KUKA KRL program: Section1.src

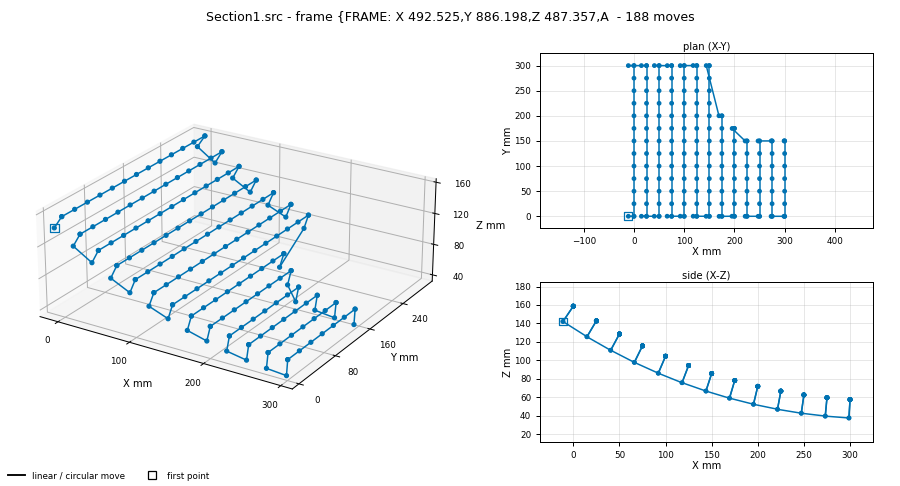
[picture p0: tool path of Section1.src in frame {FRAME: X 492.525,Y 886.198,Z 487.357,A , 188 of 189 moves have a stored position in this frame; points joined in program order, loops and branches not executed]
&ACCESS RVP
&REL 1
&PARAM TEMPLATE = C:\KRC\Roboter\Template\vorgabe
&PARAM EDITMASK = *
DEF Section1 ( )
EXT BAS (BAS_COMMAND :IN,REAL :IN )


; GLOBAL INTERRUPT DECL 3 WHEN $STOPMESS==TRUE DO IR_STOPM ( )
; INTERRUPT ON 3

;FOLD Initialise and set default speed
BAS (#INITMOV,0)
BAS (#VEL_PTP,100)
BAS (#ACC_PTP,20)
$VEL.CP=0.2
BAS (#TOOL,0)
BAS (#BASE,0)
;ENDFOLD

;;FOLD STARTPOS
;$BWDSTART = FALSE
;PDAT_ACT = PDEFAULT
;BAS(#PTP_DAT)
;FDAT_ACT = {TOOL_NO 0,BASE_NO 0,IPO_FRAME #BASE}
;BAS(#FRAMES)
;;ENDFOLD

$ADVANCE = 5

;FOLD ---- Quickly skip BCO ----
; PTP $AXIS_ACT
;ENDFOLD

;FOLD ---- GO HOME ----
; PTP {A1 0.000, A2 -90.000, A3 90.000, A4 0.000, A5 0.000, A6 0.000, E1 0, E2 0, E3 0, E4 0, E5 0, E6 0}
;ENDFOLD


; Program generated by VerticalBot Studio for KUKA KR 5 arc on 25/10/2026 12:00:00
; Using nominal kinematics.
; ---- Setting reference (Base) ----
; BASE_DATA[1] = {FRAME: X 492.525,Y 886.198,Z 487.357,A 87.824,B 90.000,C 0.000}
$BASE = {FRAME: X 492.525,Y 886.198,Z 487.357,A 87.824,B 90.000,C 0.000}
; $BASE = BASE_DATA[1]
; --------------------------
; ---- Setting tool (TCP) ----
$TOOL = {FRAME: X 25.000,Y 0.000,Z 225.000,A 0.000,B 30.000,C 0.000}
; --------------------------
; show Paint gun
$VEL.CP = 1.00000
PTP {A1 -66.38630,A2 -78.06180,A3 119.38400,A4 136.02800,A5 16.79140,A6 145.96200}
LIN {X -11.194,Y -0.005,Z 142.140,A 88.999,B 0.694,C 34.030}
LIN {X 0.000,Y 0.000,Z 158.714,A 88.999,B 0.694,C 34.030}
LIN {X 0.000,Y 0.000,Z 158.714,A 88.999,B 0.694,C 34.030}
$VEL.CP = 0.02000
LIN {X 0.000,Y 25.000,Z 158.706,A 88.999,B 0.694,C 34.030}
LIN {X 0.000,Y 50.000,Z 158.698,A 88.999,B 0.694,C 34.030}
LIN {X 0.000,Y 75.000,Z 158.689,A 88.999,B 0.695,C 34.022}
LIN {X 0.000,Y 100.000,Z 158.681,A 88.999,B 0.695,C 34.022}
LIN {X 0.000,Y 125.000,Z 158.672,A 88.999,B 0.695,C 34.022}
LIN {X 0.000,Y 150.000,Z 158.664,A 88.999,B 0.695,C 34.022}
LIN {X 0.000,Y 175.000,Z 158.655,A 88.999,B 0.695,C 34.022}
LIN {X 0.000,Y 200.000,Z 158.647,A 88.999,B 0.695,C 34.022}
LIN {X 0.000,Y 225.000,Z 158.638,A 88.999,B 0.695,C 34.022}
LIN {X 0.000,Y 250.000,Z 158.630,A 88.999,B 0.695,C 34.022}
LIN {X 0.000,Y 275.000,Z 158.628,A 88.985,B 0.696,C 34.438}
LIN {X 0.000,Y 300.000,Z 158.634,A 88.981,B 0.668,C 34.022}
$VEL.CP = 1.00000
LIN {X 0.000,Y 300.000,Z 158.634,A 88.981,B 0.668,C 34.022}
LIN {X -11.192,Y 300.006,Z 142.059,A 88.981,B 0.668,C 34.022}
$VEL.CP = 1.00000
LIN {X 14.800,Y 300.034,Z 125.622,A 88.995,B 0.482,C 30.661}
LIN {X 25.000,Y 300.000,Z 142.825,A 88.995,B 0.482,C 30.661}
LIN {X 25.000,Y 300.000,Z 142.825,A 88.995,B 0.482,C 30.661}
$VEL.CP = 0.02000
LIN {X 25.000,Y 275.000,Z 142.758,A 89.004,B 0.509,C 30.830}
LIN {X 25.000,Y 250.000,Z 142.800,A 89.264,B 0.921,C 30.374}
LIN {X 25.000,Y 225.000,Z 142.817,A 88.955,B 0.414,C 30.654}
LIN {X 25.000,Y 200.000,Z 142.818,A 89.100,B 0.691,C 31.206}
LIN {X 25.000,Y 175.000,Z 142.825,A 88.923,B 0.380,C 30.934}
LIN {X 25.000,Y 150.000,Z 142.711,A 88.930,B 0.392,C 30.935}
LIN {X 25.000,Y 125.000,Z 142.731,A 89.108,B 0.682,C 30.827}
LIN {X 25.000,Y 100.000,Z 142.834,A 88.962,B 0.476,C 31.406}
LIN {X 25.000,Y 75.000,Z 142.753,A 88.812,B 0.195,C 30.940}
LIN {X 25.000,Y 50.000,Z 142.717,A 89.127,B 0.702,C 30.616}
LIN {X 25.000,Y 25.000,Z 142.723,A 89.019,B 0.516,C 30.561}
LIN {X 25.000,Y 0.000,Z 142.733,A 88.984,B 0.455,C 30.523}
$VEL.CP = 1.00000
LIN {X 25.000,Y 0.000,Z 142.733,A 88.984,B 0.455,C 30.523}
LIN {X 14.841,Y 0.043,Z 125.505,A 88.984,B 0.455,C 30.523}
$VEL.CP = 1.00000
LIN {X 40.427,Y 0.060,Z 110.917,A 89.002,B 0.347,C 28.596}
LIN {X 50.000,Y 0.000,Z 128.477,A 89.002,B 0.347,C 28.596}
LIN {X 50.000,Y 0.000,Z 128.477,A 89.002,B 0.347,C 28.596}
$VEL.CP = 0.02000
LIN {X 50.000,Y 25.000,Z 128.477,A 89.055,B 0.450,C 28.681}
LIN {X 50.000,Y 50.000,Z 128.436,A 89.234,B 0.772,C 28.614}
LIN {X 50.000,Y 75.000,Z 128.405,A 89.097,B 0.484,C 28.082}
LIN {X 50.000,Y 100.000,Z 128.404,A 89.097,B 0.484,C 28.082}
LIN {X 50.000,Y 125.000,Z 128.414,A 89.059,B 0.414,C 28.083}
LIN {X 50.000,Y 150.000,Z 128.411,A 88.989,B 0.363,C 29.128}
LIN {X 50.000,Y 175.000,Z 128.512,A 89.007,B 0.361,C 28.667}
LIN {X 50.000,Y 200.000,Z 128.502,A 89.137,B 0.610,C 28.850}
LIN {X 50.000,Y 225.000,Z 128.556,A 88.829,B -0.037,C 27.876}
LIN {X 50.000,Y 250.000,Z 128.494,A 89.136,B 0.531,C 27.694}
LIN {X 50.000,Y 275.000,Z 128.451,A 88.924,B 0.110,C 27.503}
LIN {X 50.000,Y 300.000,Z 128.570,A 88.988,B 0.267,C 27.918}
$VEL.CP = 1.00000
LIN {X 50.000,Y 300.000,Z 128.570,A 88.988,B 0.267,C 27.918}
LIN {X 40.636,Y 300.083,Z 110.898,A 88.988,B 0.267,C 27.918}
$VEL.CP = 1.00000
LIN {X 66.337,Y 299.981,Z 97.698,A 89.173,B 0.456,C 25.664}
LIN {X 75.000,Y 300.000,Z 115.725,A 89.173,B 0.456,C 25.664}
LIN {X 75.000,Y 300.000,Z 115.725,A 89.173,B 0.456,C 25.664}
$VEL.CP = 0.02000
LIN {X 75.000,Y 275.000,Z 115.735,A 89.111,B 0.340,C 25.831}
LIN {X 75.000,Y 250.000,Z 115.738,A 89.127,B 0.361,C 25.668}
LIN {X 75.000,Y 225.000,Z 115.728,A 88.891,B -0.163,C 25.353}
LIN {X 75.000,Y 200.000,Z 115.663,A 89.159,B 0.410,C 25.464}
LIN {X 75.000,Y 175.000,Z 115.671,A 89.217,B 0.560,C 25.838}
LIN {X 75.000,Y 150.000,Z 115.708,A 89.092,B 0.311,C 25.947}
LIN {X 75.000,Y 125.000,Z 115.691,A 89.380,B 0.890,C 25.701}
LIN {X 75.000,Y 100.000,Z 115.709,A 88.958,B -0.043,C 25.137}
LIN {X 75.000,Y 75.000,Z 115.703,A 89.244,B 0.576,C 25.274}
LIN {X 75.000,Y 50.000,Z 115.702,A 89.038,B 0.250,C 26.516}
LIN {X 75.000,Y 25.000,Z 115.691,A 89.146,B 0.367,C 25.254}
LIN {X 75.000,Y 0.000,Z 115.727,A 88.965,B 0.110,C 26.587}
$VEL.CP = 1.00000
LIN {X 75.000,Y 0.000,Z 115.727,A 88.965,B 0.110,C 26.587}
LIN {X 66.050,Y 0.127,Z 97.842,A 88.965,B 0.110,C 26.587}
$VEL.CP = 1.00000
LIN {X 92.099,Y 0.138,Z 86.080,A 89.053,B -0.025,C 23.273}
LIN {X 100.000,Y 0.000,Z 104.453,A 89.053,B -0.025,C 23.273}
LIN {X 100.000,Y 0.000,Z 104.453,A 89.053,B -0.025,C 23.273}
$VEL.CP = 0.02000
LIN {X 100.000,Y 25.000,Z 104.347,A 89.212,B 0.386,C 23.749}
LIN {X 100.000,Y 50.000,Z 104.363,A 89.025,B -0.178,C 22.491}
LIN {X 100.000,Y 75.000,Z 104.359,A 89.276,B 0.496,C 23.280}
LIN {X 100.000,Y 100.000,Z 104.495,A 89.230,B 0.344,C 22.791}
LIN {X 100.000,Y 125.000,Z 104.402,A 89.329,B 0.547,C 22.387}
LIN {X 100.000,Y 150.000,Z 104.407,A 89.340,B 0.693,C 23.964}
LIN {X 100.000,Y 175.000,Z 104.463,A 89.458,B 0.826,C 21.873}
LIN {X 100.000,Y 200.000,Z 104.380,A 89.275,B 0.457,C 22.847}
LIN {X 100.000,Y 225.000,Z 104.374,A 89.143,B 0.168,C 23.111}
LIN {X 100.000,Y 250.000,Z 104.389,A 89.549,B 1.105,C 22.808}
LIN {X 100.000,Y 275.000,Z 104.335,A 89.207,B 0.310,C 23.024}
LIN {X 100.000,Y 300.000,Z 104.415,A 89.286,B 0.503,C 23.099}
$VEL.CP = 1.00000
LIN {X 100.000,Y 300.000,Z 104.415,A 89.286,B 0.503,C 23.099}
LIN {X 92.152,Y 299.936,Z 86.019,A 89.286,B 0.503,C 23.099}
$VEL.CP = 1.00000
LIN {X 117.797,Y 300.176,Z 75.721,A 89.087,B -0.188,C 21.115}
LIN {X 125.000,Y 300.000,Z 94.378,A 89.087,B -0.188,C 21.115}
LIN {X 125.000,Y 300.000,Z 94.378,A 89.087,B -0.188,C 21.115}
$VEL.CP = 0.02000
LIN {X 125.000,Y 275.000,Z 94.391,A 89.248,B 0.171,C 20.548}
LIN {X 125.000,Y 250.000,Z 94.390,A 89.138,B -0.125,C 20.520}
LIN {X 125.000,Y 225.000,Z 94.368,A 89.218,B 0.198,C 21.572}
LIN {X 125.000,Y 200.000,Z 94.368,A 89.330,B 0.321,C 19.849}
LIN {X 125.000,Y 175.000,Z 94.390,A 89.316,B 0.292,C 19.952}
LIN {X 125.000,Y 150.000,Z 94.409,A 89.332,B 0.339,C 19.984}
LIN {X 125.000,Y 125.000,Z 94.445,A 89.410,B 0.591,C 20.406}
LIN {X 125.000,Y 100.000,Z 94.434,A 89.198,B 0.012,C 20.316}
LIN {X 125.000,Y 75.000,Z 94.374,A 89.331,B 0.373,C 20.330}
LIN {X 125.000,Y 50.000,Z 94.362,A 89.240,B 0.186,C 20.895}
LIN {X 125.000,Y 25.000,Z 94.359,A 89.351,B 0.519,C 21.368}
LIN {X 125.000,Y 0.000,Z 94.453,A 89.145,B -0.084,C 20.716}
$VEL.CP = 1.00000
LIN {X 125.000,Y 0.000,Z 94.453,A 89.145,B -0.084,C 20.716}
LIN {X 117.926,Y 0.133,Z 75.746,A 89.145,B -0.084,C 20.716}
$VEL.CP = 1.00000
LIN {X 143.686,Y 0.022,Z 66.749,A 89.328,B 0.158,C 18.403}
LIN {X 150.000,Y 0.000,Z 85.726,A 89.328,B 0.158,C 18.403}
LIN {X 150.000,Y 0.000,Z 85.726,A 89.328,B 0.158,C 18.403}
$VEL.CP = 0.02000
LIN {X 150.000,Y 25.000,Z 85.716,A 89.445,B 0.525,C 18.567}
LIN {X 150.000,Y 50.000,Z 85.635,A 89.342,B 0.198,C 18.388}
LIN {X 150.000,Y 75.000,Z 85.641,A 89.365,B 0.247,C 18.195}
LIN {X 150.000,Y 100.000,Z 85.680,A 89.429,B 0.370,C 17.533}
LIN {X 150.000,Y 125.000,Z 85.656,A 89.316,B 0.069,C 17.980}
LIN {X 150.000,Y 150.000,Z 85.678,A 89.294,B 0.032,C 18.221}
LIN {X 150.000,Y 175.000,Z 85.669,A 89.401,B 0.363,C 18.285}
LIN {X 150.000,Y 200.000,Z 85.687,A 89.297,B 0.055,C 18.320}
LIN {X 150.000,Y 225.000,Z 85.698,A 89.264,B -0.104,C 17.886}
LIN {X 150.000,Y 250.000,Z 85.668,A 89.400,B 0.324,C 17.932}
LIN {X 150.000,Y 275.000,Z 85.701,A 89.532,B 0.786,C 18.614}
LIN {X 150.000,Y 300.000,Z 85.691,A 89.304,B 0.011,C 17.811}
$VEL.CP = 1.00000
LIN {X 150.000,Y 300.000,Z 85.691,A 89.304,B 0.011,C 17.811}
LIN {X 143.883,Y 300.070,Z 66.650,A 89.304,B 0.011,C 17.811}
$VEL.CP = 1.00000
LIN {X 169.191,Y 200.159,Z 59.012,A 89.262,B -0.253,C 16.891}
LIN {X 175.000,Y 200.000,Z 78.149,A 89.262,B -0.253,C 16.891}
LIN {X 175.000,Y 200.000,Z 78.149,A 89.262,B -0.253,C 16.891}
$VEL.CP = 0.02000
LIN {X 175.000,Y 175.000,Z 78.173,A 89.333,B -0.189,C 15.738}
LIN {X 175.000,Y 150.000,Z 78.128,A 89.417,B 0.046,C 15.303}
LIN {X 175.000,Y 125.000,Z 78.138,A 89.425,B 0.132,C 15.692}
LIN {X 175.000,Y 100.000,Z 78.159,A 89.394,B 0.073,C 16.078}
LIN {X 175.000,Y 75.000,Z 78.141,A 89.431,B 0.093,C 15.272}
LIN {X 175.000,Y 50.000,Z 78.135,A 89.438,B 0.177,C 15.711}
LIN {X 175.000,Y 25.000,Z 78.230,A 89.557,B 0.606,C 15.756}
LIN {X 175.000,Y 0.000,Z 78.195,A 89.528,B 0.537,C 16.065}
$VEL.CP = 1.00000
LIN {X 175.000,Y 0.000,Z 78.195,A 89.528,B 0.537,C 16.065}
LIN {X 169.464,Y -0.134,Z 58.977,A 89.528,B 0.537,C 16.065}
$VEL.CP = 1.00000
LIN {X 195.189,Y 0.101,Z 52.416,A 89.422,B -0.156,C 13.921}
LIN {X 200.000,Y 0.000,Z 71.829,A 89.422,B -0.156,C 13.921}
LIN {X 200.000,Y 0.000,Z 71.829,A 89.422,B -0.156,C 13.921}
$VEL.CP = 0.02000
LIN {X 200.000,Y 25.000,Z 71.844,A 89.490,B 0.058,C 13.542}
LIN {X 200.000,Y 50.000,Z 71.795,A 89.530,B 0.139,C 12.980}
LIN {X 200.000,Y 75.000,Z 71.810,A 89.522,B 0.096,C 12.941}
LIN {X 200.000,Y 100.000,Z 71.796,A 89.527,B 0.125,C 12.978}
LIN {X 200.000,Y 125.000,Z 71.872,A 89.573,B 0.354,C 13.177}
LIN {X 200.000,Y 150.000,Z 71.817,A 89.505,B -0.092,C 12.310}
LIN {X 200.000,Y 175.000,Z 71.807,A 89.602,B 0.473,C 13.157}
$VEL.CP = 1.00000
LIN {X 200.000,Y 175.000,Z 71.807,A 89.602,B 0.473,C 13.157}
LIN {X 195.447,Y 174.871,Z 52.332,A 89.602,B 0.473,C 13.157}
$VEL.CP = 1.00000
LIN {X 221.328,Y 149.942,Z 46.992,A 89.638,B 0.237,C 10.579}
LIN {X 225.000,Y 150.000,Z 66.652,A 89.638,B 0.237,C 10.579}
LIN {X 225.000,Y 150.000,Z 66.652,A 89.638,B 0.237,C 10.579}
$VEL.CP = 0.02000
LIN {X 225.000,Y 125.000,Z 66.645,A 89.661,B 0.444,C 11.059}
LIN {X 225.000,Y 100.000,Z 66.702,A 89.684,B 0.470,C 10.495}
LIN {X 225.000,Y 75.000,Z 66.641,A 89.560,B -0.271,C 10.190}
LIN {X 225.000,Y 50.000,Z 66.583,A 89.646,B 0.139,C 9.851}
LIN {X 225.000,Y 25.000,Z 66.619,A 89.653,B 0.483,C 11.578}
LIN {X 225.000,Y 0.000,Z 66.575,A 89.608,B 0.035,C 10.373}
$VEL.CP = 1.00000
LIN {X 225.000,Y 0.000,Z 66.575,A 89.608,B 0.035,C 10.373}
LIN {X 221.399,Y 0.013,Z 46.902,A 89.608,B 0.035,C 10.373}
$VEL.CP = 1.00000
LIN {X 247.259,Y -0.014,Z 42.649,A 89.710,B 0.081,C 7.876}
LIN {X 250.000,Y 0.000,Z 62.461,A 89.710,B 0.081,C 7.876}
LIN {X 250.000,Y 0.000,Z 62.461,A 89.710,B 0.081,C 7.876}
$VEL.CP = 0.02000
LIN {X 250.000,Y 25.000,Z 62.499,A 89.666,B -0.292,C 7.715}
LIN {X 250.000,Y 50.000,Z 62.506,A 89.689,B 0.029,C 8.245}
LIN {X 250.000,Y 75.000,Z 62.507,A 89.697,B 0.077,C 8.213}
LIN {X 250.000,Y 100.000,Z 62.503,A 89.732,B 0.235,C 7.860}
LIN {X 250.000,Y 125.000,Z 62.545,A 89.664,B -0.225,C 7.962}
LIN {X 250.000,Y 150.000,Z 62.456,A 89.683,B 0.028,C 8.391}
$VEL.CP = 1.00000
LIN {X 250.000,Y 150.000,Z 62.456,A 89.683,B 0.028,C 8.391}
LIN {X 247.081,Y 150.006,Z 42.670,A 89.683,B 0.028,C 8.391}
$VEL.CP = 1.00000
LIN {X 273.289,Y 150.082,Z 39.572,A 89.794,B -0.219,C 4.909}
LIN {X 275.000,Y 150.000,Z 59.499,A 89.794,B -0.219,C 4.909}
LIN {X 275.000,Y 150.000,Z 59.499,A 89.794,B -0.219,C 4.909}
$VEL.CP = 0.02000
LIN {X 275.000,Y 125.000,Z 59.428,A 89.772,B 0.109,C 6.284}
LIN {X 275.000,Y 100.000,Z 59.496,A 89.797,B -0.199,C 4.874}
LIN {X 275.000,Y 75.000,Z 59.566,A 89.798,B 0.309,C 6.164}
LIN {X 275.000,Y 50.000,Z 59.574,A 89.738,B -0.250,C 6.168}
LIN {X 275.000,Y 25.000,Z 59.452,A 89.738,B -0.250,C 6.168}
LIN {X 275.000,Y 0.000,Z 59.424,A 89.789,B 0.061,C 5.689}
$VEL.CP = 1.00000
LIN {X 275.000,Y 0.000,Z 59.424,A 89.789,B 0.061,C 5.689}
LIN {X 273.017,Y -0.014,Z 39.523,A 89.789,B 0.061,C 5.689}
$VEL.CP = 1.00000
LIN {X 298.681,Y -0.024,Z 37.514,A 89.861,B 0.079,C 3.780}
LIN {X 300.000,Y 0.000,Z 57.470,A 89.861,B 0.079,C 3.780}
LIN {X 300.000,Y 0.000,Z 57.470,A 89.861,B 0.079,C 3.780}
$VEL.CP = 0.02000
LIN {X 300.000,Y 25.000,Z 57.480,A 89.885,B 0.092,C 3.162}
LIN {X 300.000,Y 50.000,Z 57.449,A 89.852,B -0.049,C 3.801}
LIN {X 300.000,Y 75.000,Z 57.506,A 89.843,B -0.185,C 3.800}
LIN {X 300.000,Y 100.000,Z 57.488,A 89.901,B 0.252,C 2.944}
LIN {X 300.000,Y 125.000,Z 57.438,A 89.871,B -0.047,C 3.316}
LIN {X 300.000,Y 150.000,Z 57.492,A 89.860,B -0.386,C 3.131}
$VEL.CP = 1.00000
LIN {X 300.000,Y 150.000,Z 57.492,A 89.860,B -0.386,C 3.131}
LIN {X 298.908,Y 150.137,Z 37.523,A 89.860,B -0.386,C 3.131}
END
